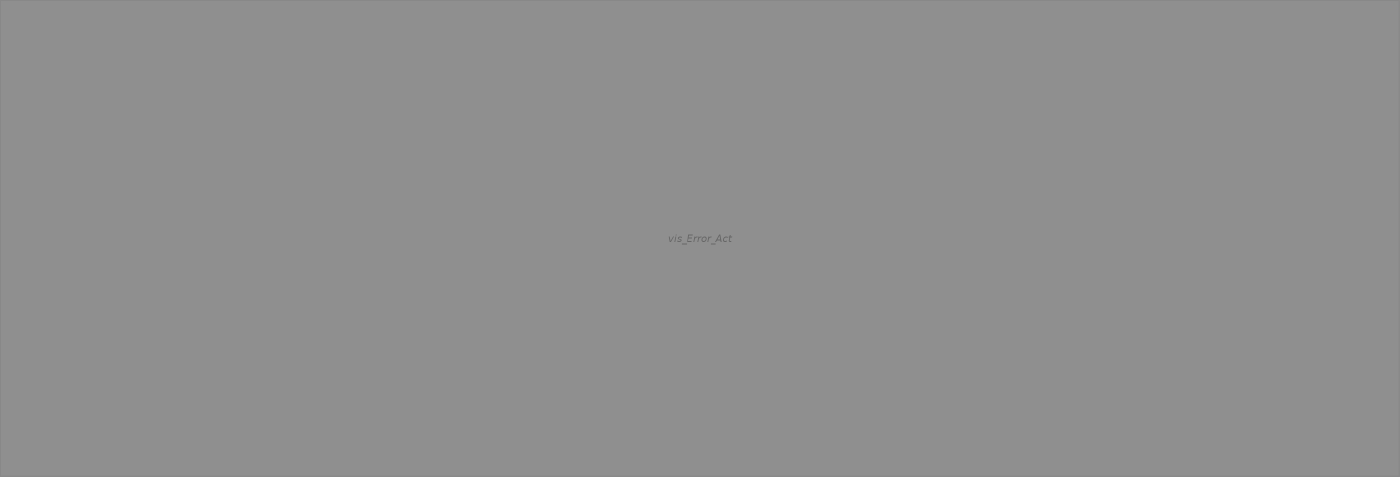
VISUALIZATION ERROR_Tab  // 1428x487
    Rectangle (0,0 1428x487)
    TabControl (0,0 1428x487)
        shows vis_Error_Act()
        shows vis_Error_History()
        shows vis_Error_Search()
        [0]: TabTitle=Actual Errors
        [1]: TabTitle=Error History
        [2]: TabTitle=Search
END_VISUALIZATION

(* stored: Version 1.1.0.1, ProductVersion 3.1.4024.13
   Visu ERROR_Tab: Id {12037b74-6a44-40c8-8fc7-653dfd555b55} *)
